// TIA Portal V20 export
ScreenOverview   800x60
  ScreenLayer 
    SymbolicIOField "Symbolic_IO_Field_Screen" at 109,11 size 584x38  CountVisibleItems=3, Mode=InOutput, OnValue=1, TextList=TextList_ScreenNames, TextOff="0", TextOn="1"
      on Change: ActivateScreenByNumber(Screen number := Tag_ScreenNumber, Object number := 0)
      ProcessValue := Tag_ScreenNumber
    DateTimeField "HmiScreenItemData" at 695,30 size 105x30  Mode=Output
    DateTimeField "HmiScreenItemData_1" at 695,0 size 105x30  Mode=Output
    GraphicView "Logo" at 0,0 size 107x60  Picture=Logo of HMI_1
